(* Status of spindle *)

TYPE ET_SpindleClutchStatus :
(
	ET_SpindleClutchStatus_ClosedWithoutTool := 0,				(* Clutch is closed without tool *)
	ET_SpindleClutchStatus_ClosedWithTool := 1,					(* Clutch is closed with tool *)
	ET_SpindleClutchStatus_Opened := 2,						(* Clutch is opened *)
	ET_SpindleClutchStatus_RotatingNoClosed := 3,				(* Clutch rotating and not closed *)
	ET_SpindleClutchStatus_NoDefined := 999
);
END_TYPE

(* stored: Version 1.1.0.1, ProductVersion 3.1.4024.15
   DUT ET_SpindleClutchStatus: Id {91da0715-b0c1-4d3b-a018-b88339286977} *)
